(* IEC 61131-3 sources: trust-platform/editors/vscode/src/test/fixtures/control-studio-two-zone-group/src, 1 file *)

(* ---- Main.st ---- *)
USING Control;

(* Two heated zones that share a wall, one Control.PID per zone and one Auto/Manual switch for both, so the
   two controllers are commissioned together as a group. Heating one zone also warms the other. *)
PROGRAM Main
VAR
    Zone1 : Control.PID;
    Zone2 : Control.PID;
    Zone1Parameters : Control.PIDParameters := (
        ProportionalGain := LREAL#4.0, IntegralGain := LREAL#0.5, DerivativeGain := LREAL#0.0,
        ProportionalSetpointWeight := LREAL#1.0, DerivativeSetpointWeight := LREAL#0.0, Bias := LREAL#0.0,
        OutputMinimum := LREAL#0.0, OutputMaximum := LREAL#100.0,
        RateMinimum := LREAL#-1000.0, RateMaximum := LREAL#1000.0, TrackingTime := LREAL#1.0,
        AntiWindup := PIDAntiWindup#BackCalculation);
    Zone2Parameters : Control.PIDParameters := (
        ProportionalGain := LREAL#4.0, IntegralGain := LREAL#0.5, DerivativeGain := LREAL#0.0,
        ProportionalSetpointWeight := LREAL#1.0, DerivativeSetpointWeight := LREAL#0.0, Bias := LREAL#0.0,
        OutputMinimum := LREAL#0.0, OutputMaximum := LREAL#100.0,
        RateMinimum := LREAL#-1000.0, RateMaximum := LREAL#1000.0, TrackingTime := LREAL#1.0,
        AntiWindup := PIDAntiWindup#BackCalculation);
    Zone1Input : Control.PIDInput;
    Zone2Input : Control.PIDInput;
    State : Control.PIDInitialState;
    Initialized : BOOL := FALSE;
    (* TRUE selects Auto for both controllers; they start in Manual at the resting point. *)
    ZonesAuto : BOOL := FALSE;
    Zone1ManualPct : LREAL := 20.0;
    Zone2ManualPct : LREAL := 20.0;
    Zone1SetpointC : LREAL := 26.0;
    Zone2SetpointC : LREAL := 26.0;
    Zone1C : LREAL := 26.0;
    Zone2C : LREAL := 26.0;
    Heater1Pct : LREAL := 20.0;
    Heater2Pct : LREAL := 20.0;
END_VAR

Zone1.Configure(Parameters := Zone1Parameters);
Zone2.Configure(Parameters := Zone2Parameters);
IF NOT Initialized THEN
    (* Memory-mapped variables start from the %M image; set the resting values explicitly. *)
    Zone1SetpointC := LREAL#26.0;
    Zone2SetpointC := LREAL#26.0;
    Zone1ManualPct := LREAL#20.0;
    Zone2ManualPct := LREAL#20.0;
    State.Setpoint := Zone1SetpointC;
    State.ProcessValue := Zone1C;
    State.NominalOutput := Zone1ManualPct;
    State.SaturatedOutput := Zone1ManualPct;
    Zone1.Initialize(State := State);
    State.Setpoint := Zone2SetpointC;
    State.ProcessValue := Zone2C;
    State.NominalOutput := Zone2ManualPct;
    State.SaturatedOutput := Zone2ManualPct;
    Zone2.Initialize(State := State);
    Initialized := TRUE;
END_IF;

Zone1Input.Setpoint := Zone1SetpointC;
Zone1Input.ProcessValue := Zone1C;
Zone1Input.ManualOutput := Zone1ManualPct;
Zone1Input.TrackingOutput := Zone1ManualPct;
Zone1Input.CycleTime := LREAL#0.1;
IF ZonesAuto THEN
    Zone1Input.Mode := PIDMode#Auto;
ELSE
    Zone1Input.Mode := PIDMode#Manual;
END_IF;
Heater1Pct := Zone1.Update(Input := Zone1Input);

Zone2Input.Setpoint := Zone2SetpointC;
Zone2Input.ProcessValue := Zone2C;
Zone2Input.ManualOutput := Zone2ManualPct;
Zone2Input.TrackingOutput := Zone2ManualPct;
Zone2Input.CycleTime := LREAL#0.1;
IF ZonesAuto THEN
    Zone2Input.Mode := PIDMode#Auto;
ELSE
    Zone2Input.Mode := PIDMode#Manual;
END_IF;
Heater2Pct := Zone2.Update(Input := Zone2Input);
END_PROGRAM

CONFIGURATION Config
RESOURCE Res ON PLC
    TASK MainTask(INTERVAL := T#100ms, PRIORITY := 1);
    PROGRAM P1 WITH MainTask : Main;
END_RESOURCE
VAR_CONFIG
    P1.Heater1Pct AT %QL0 : LREAL;
    P1.Heater2Pct AT %QL8 : LREAL;
    P1.Zone1C AT %IL0 : LREAL;
    P1.Zone2C AT %IL8 : LREAL;
    P1.Zone1SetpointC AT %ML0 : LREAL;
    P1.Zone2SetpointC AT %ML8 : LREAL;
    P1.Zone1ManualPct AT %ML16 : LREAL;
    P1.Zone2ManualPct AT %ML24 : LREAL;
END_VAR
END_CONFIGURATION
